FUNCTION_BLOCK FB_ControlPanel
VAR_INPUT
	bStartPB    : BOOL;  // physical start, NO (TRUE = pressed)
	bStopPB     : BOOL;  // physical stop, NC (FALSE = pressed)
	bEStopPB    : BOOL;  // physical emergency, NC (FALSE = pressed)
	bHmiStart   : BOOL;  // soft buttons from HMI
	bHmiStop    : BOOL;
	bHmiEStop   : BOOL;
	bReset      : BOOL;  // felles reset (HMI)
END_VAR
VAR_OUTPUT
	bRunning    : BOOL;  // process is allowed to run
	bEmergency  : BOOL;  // latched emergency, needs reset
	bStopActive : BOOL;  // a stop is being requested right now
END_VAR
VAR
	rtStart     : R_TRIG;
	rtHmiStart  : R_TRIG;
END_VAR

// Flankedeteksjon på start
rtStart(CLK := bStartPB);
rtHmiStart(CLK := bHmiStart);

// Stopp = fysisk NC åpnet ELLER soft stop (inkl. trip fra MAIN)
bStopActive := NOT bStopPB OR bHmiStop;

// Nødstopp låses. Kvitteres kun med bReset når nødstoppen er sluppet
IF NOT bEStopPB OR bHmiEStop THEN
	bEmergency := TRUE;
ELSIF bEmergency AND bReset THEN
	bEmergency := FALSE;
END_IF

// Start på stigende flanke, kun når ingen stopp eller nødstopp er aktiv
IF bEmergency OR bStopActive THEN
	bRunning := FALSE;
ELSIF rtStart.Q OR rtHmiStart.Q THEN
	bRunning := TRUE;
END_IF

END_FUNCTION_BLOCK

(* stored: Version 1.1.0.1, ProductVersion 3.1.4026.21
   POU FB_ControlPanel: Id {9efcfb52-dadb-41f6-9abe-218aa7d971fa}, SpecialFunc None *)
